// TEST DI FB_Timer
FUNCTION_BLOCK FB_Timer_Test EXTENDS TcUnit.FB_TestSuite
VAR
	fbElapsed	:	ML.FB_Timer;
	fbSelf		:	ML.FB_Timer;
	fbReset		:	ML.FB_Timer;
END_VAR

VerifyElapsed();
VerifySelfElapsed();
ResetCondition();

METHOD PRIVATE ResetCondition
TEST('ResetCondition');

fbReset.ResetWithOffset(T#5S);
AssertFalse(Condition := fbReset.ResetCondition(FALSE),	Message := 'Condizione FALSE: nessun reset');
AssertTrue(Condition := fbReset.VerifyElapsed(T#4S),		Message := 'Senza reset il tempo trascorso resta 5 s');
AssertTrue(Condition := fbReset.ResetCondition(TRUE),		Message := 'Condizione TRUE: reset eseguito');
AssertFalse(Condition := fbReset.VerifyElapsed(T#1S),		Message := 'Dopo il reset il tempo riparte da 0');

TEST_FINISHED();
END_METHOD

METHOD PRIVATE VerifyElapsed
TEST('VerifyElapsed');

fbElapsed.ResetWithOffset(T#2S);
AssertTrue(Condition := fbElapsed.VerifyElapsed(T#1S),	Message := 'Sono passati 2 s: 1 s deve risultare trascorso');
AssertFalse(Condition := fbElapsed.VerifyElapsed(T#10S),	Message := 'Sono passati 2 s: 10 s non devono risultare trascorsi');

TEST_FINISHED();
END_METHOD

METHOD PRIVATE VerifySelfElapsed
TEST('VerifySelfElapsed');

fbSelf.ResetWithOffset(T#2S);
fbSelf.ChangeTimer(T#1S);
AssertTrue(Condition := fbSelf.VerifySelfElapsed(),	Message := 'Durata 1 s, trascorsi 2 s');
fbSelf.ChangeTimer(T#10S);
AssertFalse(Condition := fbSelf.VerifySelfElapsed(),	Message := 'Durata 10 s, trascorsi 2 s');

TEST_FINISHED();
END_METHOD

END_FUNCTION_BLOCK

(* stored: Version 1.1.0.1, ProductVersion 3.1.4024.9
   POU FB_Timer_Test: Id {c74504a1-f754-4e83-a888-25eac838705e}, SpecialFunc None
   Folder METHODs: Id {5ce43d5c-5da5-45c1-a934-98a1346bfd4f}
   Method ResetCondition: Id {a2714dce-b0c1-452a-bec5-7a3f58e3825d}
   Method VerifyElapsed: Id {0aa4564d-23e8-4f55-a3cc-fe4d3601d0c0}
   Method VerifySelfElapsed: Id {0e1758b8-3b8d-40f6-ab70-ec4d2cb5b193} *)
